Universal Robots URScript: T002_openai_gpt-oss-120b_baseline_rep1.urscript

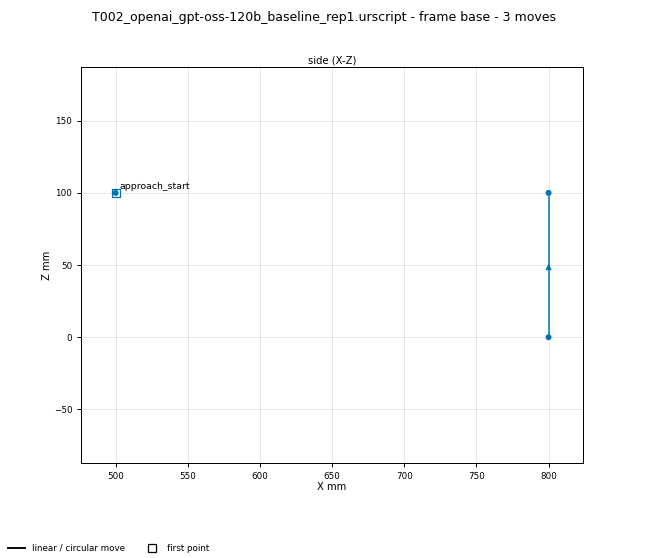
[picture p0: tool path of T002_openai_gpt-oss-120b_baseline_rep1.urscript in frame base, 3 of 6 moves have a stored position in this frame; points joined in program order, loops and branches not executed]
def main():
    # -------------------------------------------------
    # Configuration
    # -------------------------------------------------
    # Payload
    set_payload(3.0, [0, 0, 0.1])          # 3 kg, CoG 10 cm above TCP

    # Tool (placeholder, 20 mm length)
    set_tcp([0, 0, 0.02, 0, 0, 0])

    # Safety: fenced (confinement & exclusion zones)
    set_fence_enabled(True)                # Enable fenced mode
    # (Optional: define explicit zones if required)
    # set_confinement_zone([[0.3, -0.3, 0.0, 0.0, 0.0, 0.0], [1.0, 0.3, 0.5, 0.0, 0.0, 0.0]])
    # set_exclusion_zone([[0.0, -0.2, 0.0, 0.0, 0.0, 0.0], [0.2, 0.2, 0.5, 0.0, 0.0, 0.0]])

    # -------------------------------------------------
    # Pose definitions (meters, radians)
    # -------------------------------------------------
    # Home joint configuration (UR5e default)
    home_joints = [-0.0, -1.5708, 1.5708, -1.5708, -1.5708, 0.0]

    # Weld start (on workpiece surface)
    weld_start = p[0.500, 0.000, 0.000, 0.0, 3.14159, 0.0]   # orientation: torch pointing down

    # Approach point 10 cm above start
    approach_start = p[0.500, 0.000, 0.100, 0.0, 3.14159, 0.0]

    # Weld end (300 mm along X)
    weld_end = p[0.800, 0.000, 0.000, 0.0, 3.14159, 0.0]

    # Retract point 10 cm above end
    retract_end = p[0.800, 0.000, 0.100, 0.0, 3.14159, 0.0]

    # -------------------------------------------------
    # Motion sequence
    # -------------------------------------------------
    # 1) Move to home position
    movej(home_joints, a=1.2, v=0.300)   # 300 mm/s

    # 2) Approach above weld start
    movel(approach_start, a=1.2, v=0.250)   # 250 mm/s

    # 3) Descend to weld start position
    movel(weld_start, a=1.2, v=0.100)       # 100 mm/s

    # 4) Activate welding (digital output 0)
    set_digital_out(0, True)

    # 5) Weld seam – 300 mm linear path
    #    Speed limited to 50 mm/s for welding arc
    movel(weld_end, a=0.5, v=0.050)         # 50 mm/s

    # 6) Deactivate welding
    set_digital_out(0, False)

    # 7) Retract above weld end
    movel(retract_end, a=1.2, v=0.200)      # 200 mm/s

    # 8) Return to home position
    movej(home_joints, a=1.2, v=0.300)

    # -------------------------------------------------
    # End of program
    # -------------------------------------------------
    set_fence_enabled(False)   # Disable fenced mode (optional)
end

# -----------------------------------------------------------------
# Run the program
# -----------------------------------------------------------------
main()
